(* IEC 61131-3 sources: JingjiangMoonbox/Application/Application/任务列表/CommTask/参数初始化 (part 2) *)

(* ---- KS_RstGrpParam_UnSave.st ---- *)
(*@CES
Name=KS_RstGrpParam_UnSave
Type=FunctionBlock
TypeGuid=6f9dac99-8de1-4efc-8465-68ac443b7d08
Guid=192eb973-c984-42d3-866b-81e626ce7a5f
HasDeclaration=True
HasImplementation=True
*)
{DECLARATION}
FUNCTION KS_RstGrpParam_UnSave : INT
VAR_INPUT
	i_pastStGrpParam_UnSave: POINTER TO ARRAY [1..2] OF StGrpParam_UnSave;
	i_pastStGrpParam_UnSave_RSV: POINTER TO ARRAY [1..2] OF StRSV_GrpParam_UnSave;
END_VAR
VAR
	iGrp: INT;
	iResult: INT;
	iT: INT;
END_VAR

{IMPLEMENTATION}
iResult:=0;

IF i_pastStGrpParam_UnSave<>0 AND i_pastStGrpParam_UnSave_RSV<>0 THEN
	FOR iGrp:=1 TO 2 BY 1 DO
		SysMemSet(ADR(i_pastStGrpParam_UnSave_RSV^[iGrp].abyRSV_StGrpParam_UnSave),
					0,
					SIZEOF(i_pastStGrpParam_UnSave_RSV^[iGrp].abyRSV_StGrpParam_UnSave));
		i_pastStGrpParam_UnSave^[iGrp].xCutterOnTop_Uw						:= TRUE;
		i_pastStGrpParam_UnSave^[iGrp].iDebugVelmpm_AxisA_Uw                := 100;
		i_pastStGrpParam_UnSave^[iGrp].iDebugGirthmm_AxisA_Uw               := 300;
		i_pastStGrpParam_UnSave^[iGrp].iDebugVelmpm_AxisB_Uw                := 100;
		i_pastStGrpParam_UnSave^[iGrp].iDebugGirthmm_AxisB_Uw               := 300;
		i_pastStGrpParam_UnSave^[iGrp].iDebugVelmpm_AxisA_Rw                := 100;
		i_pastStGrpParam_UnSave^[iGrp].iDebugGirthmm_AxisA_Rw               := 300;
		i_pastStGrpParam_UnSave^[iGrp].iDebugVelmpm_AxisB_Rw                := 100;
		i_pastStGrpParam_UnSave^[iGrp].iDebugGirthmm_AxisB_Rw               := 300;
		i_pastStGrpParam_UnSave^[iGrp].xMachineRev                          := FALSE;
		i_pastStGrpParam_UnSave^[iGrp].iPromptMsg                           := 0;
		i_pastStGrpParam_UnSave^[iGrp].iAlarm_TypeId                        := 0;
		i_pastStGrpParam_UnSave^[iGrp].iAlarm_UnitId                        := 0;
		i_pastStGrpParam_UnSave^[iGrp].iIdGSE                               := GSE_STOP;
		i_pastStGrpParam_UnSave^[iGrp].xFlag_Stop                           := TRUE;
		i_pastStGrpParam_UnSave^[iGrp].xFlag_PreStart                       := FALSE;
		i_pastStGrpParam_UnSave^[iGrp].xFlag_Ink                            := FALSE;
		i_pastStGrpParam_UnSave^[iGrp].xFlag_InkAccing                      := FALSE;
		i_pastStGrpParam_UnSave^[iGrp].xFlag_Tension                        := FALSE;
		i_pastStGrpParam_UnSave^[iGrp].xFlag_TensionDone                    := FALSE;
		i_pastStGrpParam_UnSave^[iGrp].xFlag_Print                          := FALSE;
		i_pastStGrpParam_UnSave^[iGrp].xFlag_Estop                          := FALSE;
		i_pastStGrpParam_UnSave^[iGrp].xFlag_AutoAcc                        := FALSE;
		i_pastStGrpParam_UnSave^[iGrp].xFlag_AutoDec                        := FALSE;
		i_pastStGrpParam_UnSave^[iGrp].xFlag_ManuAcc                        := FALSE;
		i_pastStGrpParam_UnSave^[iGrp].xFlag_ManuDec                        := FALSE;
		i_pastStGrpParam_UnSave^[iGrp].xFlag_Accing                         := FALSE;
		i_pastStGrpParam_UnSave^[iGrp].xFlag_Decing                         := FALSE;
		i_pastStGrpParam_UnSave^[iGrp].xFlag_EStoping                       := FALSE;
		i_pastStGrpParam_UnSave^[iGrp].xFlag_Stoping                        := FALSE;
		i_pastStGrpParam_UnSave^[iGrp].xFlag_GotoInking                     := FALSE;
		i_pastStGrpParam_UnSave^[iGrp].xFlag_InPressing                     := FALSE;
		i_pastStGrpParam_UnSave^[iGrp].xFlag_RollerPressDone                := FALSE;
		i_pastStGrpParam_UnSave^[iGrp].xFlag_InchRun                        := FALSE;
		i_pastStGrpParam_UnSave^[iGrp].xFlag_AllInchRun                     := FALSE;
		i_pastStGrpParam_UnSave^[iGrp].xFlag_AllPress                       := FALSE;
		i_pastStGrpParam_UnSave^[iGrp].xFlag_AllUnpress                     := FALSE;
		i_pastStGrpParam_UnSave^[iGrp].xFlag_RollerPressAtLeast1            := FALSE;
		i_pastStGrpParam_UnSave^[iGrp].axFlag_PrnLen_Alarm[1]                  := FALSE;
		i_pastStGrpParam_UnSave^[iGrp].axFlag_PrnLen_Alarm[2]                  := FALSE;
		i_pastStGrpParam_UnSave^[iGrp].axFlag_PrnLen_Alarm[3]                  := FALSE;
		i_pastStGrpParam_UnSave^[iGrp].xFlag_LinkageAxisAlarm               := FALSE;
		i_pastStGrpParam_UnSave^[iGrp].xFlag_TensionUnfinished              := FALSE;
		i_pastStGrpParam_UnSave^[iGrp].xFlag_VelTooHigh                     := FALSE;
		i_pastStGrpParam_UnSave^[iGrp].xFlag_PrestartTimeout                := FALSE;
		i_pastStGrpParam_UnSave^[iGrp].xFlag_KeepAlarming                   := FALSE;
		i_pastStGrpParam_UnSave^[iGrp].xFlag_ArrivedToTargetVel             := FALSE;
		i_pastStGrpParam_UnSave^[iGrp].xFlag_FilmAccDecDone                 := FALSE;
		i_pastStGrpParam_UnSave^[iGrp].xSlowStopTenEn                       := FALSE;
		i_pastStGrpParam_UnSave^[iGrp].xIsDebugMode_Machine                 := FALSE;
		i_pastStGrpParam_UnSave^[iGrp].uiFilmThickNess                      := 20;
		i_pastStGrpParam_UnSave^[iGrp].abyClrPrnLenCount_Rw[1]                 := 0;
		i_pastStGrpParam_UnSave^[iGrp].abyClrPrnLenCount_Rw[2]                 := 0;
		i_pastStGrpParam_UnSave^[iGrp].abyClrPrnLenCount_Rw[3]                 := 0;
		i_pastStGrpParam_UnSave^[iGrp].iTimeSec_AccDec_AllTheWay            := 0;
		i_pastStGrpParam_UnSave^[iGrp].rAccDecTime_ThisTime                 := 0;
		i_pastStGrpParam_UnSave^[iGrp].alrStdVol_Diam_Axis_Hmi[1]              := 0;
		i_pastStGrpParam_UnSave^[iGrp].alrStdVol_Diam_Axis_Hmi[2]              := 0;
		i_pastStGrpParam_UnSave^[iGrp].alrStdVol_Diam_Axis_Hmi[3]              := 0;
		i_pastStGrpParam_UnSave^[iGrp].alrStdVol_Diam_Axis_Hmi[4]              := 0;
		i_pastStGrpParam_UnSave^[iGrp].alrStdVol_Volt_Axis_Hmi[1]              := 0;
		i_pastStGrpParam_UnSave^[iGrp].alrStdVol_Volt_Axis_Hmi[2]              := 0;
		i_pastStGrpParam_UnSave^[iGrp].alrStdVol_Volt_Axis_Hmi[3]              := 0;
		i_pastStGrpParam_UnSave^[iGrp].alrStdVol_Volt_Axis_Hmi[4]              := 0;
		i_pastStGrpParam_UnSave^[iGrp].alrStdVol_Coef_Axis_Hmi[0]              := 0;
		i_pastStGrpParam_UnSave^[iGrp].alrStdVol_Coef_Axis_Hmi[1]              := 0;
		i_pastStGrpParam_UnSave^[iGrp].alrStdVol_Coef_Axis_Hmi[2]              := 0;
		i_pastStGrpParam_UnSave^[iGrp].alrStdVol_Coef_Axis_Hmi[3]              := 0;
		i_pastStGrpParam_UnSave^[iGrp].alrStdVol_Coef_Axis_Hmi[4]              := 0;
		i_pastStGrpParam_UnSave^[iGrp].rVel_Cur                             := 0;
		i_pastStGrpParam_UnSave^[iGrp].rVel_Film                            := 0;
		i_pastStGrpParam_UnSave^[iGrp].iSid_AxisA_Uw                        := 112;
		i_pastStGrpParam_UnSave^[iGrp].xStationOnline_AxisA_Uw              := FALSE;
		i_pastStGrpParam_UnSave^[iGrp].xMotRev_AxisA_Uw                     := FALSE;
		i_pastStGrpParam_UnSave^[iGrp].iSid_AxisB_Uw                        := 113;
		i_pastStGrpParam_UnSave^[iGrp].xStationOnline_AxisB_Uw              := FALSE;
		i_pastStGrpParam_UnSave^[iGrp].xMotRev_AxisB_Uw                     := FALSE;
		i_pastStGrpParam_UnSave^[iGrp].rAI_Uw                               := 0;
		i_pastStGrpParam_UnSave^[iGrp].rAI_Act_Uw                           := 0;
		i_pastStGrpParam_UnSave^[iGrp].rAI_HMI_Uw                           := 0;
		i_pastStGrpParam_UnSave^[iGrp].rAI_DiamMeasure_Uw                   := 0;
		i_pastStGrpParam_UnSave^[iGrp].arKpid_Current_Uw[1]                    := 20;
		i_pastStGrpParam_UnSave^[iGrp].arKpid_Current_Uw[2]                    := 50;
		i_pastStGrpParam_UnSave^[iGrp].arKpid_Current_Uw[3]                    := 50;
		i_pastStGrpParam_UnSave^[iGrp].arKpid_Current_Rw[1]                    := 0;
		i_pastStGrpParam_UnSave^[iGrp].arKpid_Current_Rw[2]                    := 0;
		i_pastStGrpParam_UnSave^[iGrp].arKpid_Current_Rw[3]                    := 0;
		i_pastStGrpParam_UnSave^[iGrp].rVel_PreDrv_Uw                       := 0;
		i_pastStGrpParam_UnSave^[iGrp].xReflectionSensorValid_Uw            := FALSE;
		i_pastStGrpParam_UnSave^[iGrp].xReflectSensorLoss_Uw                := FALSE;
		i_pastStGrpParam_UnSave^[iGrp].rDiam_NewVol_Uw                      := 400;
		i_pastStGrpParam_UnSave^[iGrp].rTowerThetaCur_Uw                    := 0;
		i_pastStGrpParam_UnSave^[iGrp].rFilmToTowerRollerDis_Uw             := 0;
		i_pastStGrpParam_UnSave^[iGrp].xFilmTouchRoller_Uw                  := FALSE;
		i_pastStGrpParam_UnSave^[iGrp].xSts_PreCutting_Uw                   := FALSE;
		i_pastStGrpParam_UnSave^[iGrp].rDebugCurVelmpmAxisA_Uw              := 0;
		i_pastStGrpParam_UnSave^[iGrp].rDebugCurVelrpmAxisA_Uw              := 0;
		i_pastStGrpParam_UnSave^[iGrp].rDebugCurVelmpmAxisB_Uw              := 0;
		i_pastStGrpParam_UnSave^[iGrp].rDebugCurVelrpmAxisB_Uw              := 0;
		i_pastStGrpParam_UnSave^[iGrp].rDeltaW_RPMIN_Uw                     := 0;
		i_pastStGrpParam_UnSave^[iGrp].xDebugMode_AbsEnc_Uw                 := FALSE;
		i_pastStGrpParam_UnSave^[iGrp].dwAbsEncSinglePos_Uw                 := 0;
		i_pastStGrpParam_UnSave^[iGrp].dwAbsEncSPos_Cur_Uw                  := 0;
		i_pastStGrpParam_UnSave^[iGrp].byEncodeValueWr_Uw                   := 0;
		i_pastStGrpParam_UnSave^[iGrp].rAIByAbsEnc_Cur_Uw                   := 0;
		i_pastStGrpParam_UnSave^[iGrp].xCutterOnTopFroDebug_Uw              := FALSE;
		i_pastStGrpParam_UnSave^[iGrp].xCurAxisAFroDebug_Uw                 := FALSE;
		i_pastStGrpParam_UnSave^[iGrp].xAlarmBell_Uw                        := FALSE;
		i_pastStGrpParam_UnSave^[iGrp].xIsDebug_DiaMeasure_Uw               := FALSE;
		i_pastStGrpParam_UnSave^[iGrp].byIsDebug_DiaMeasureArea_Uw          := 0;
		i_pastStGrpParam_UnSave^[iGrp].xIsDebuging_DiaMeasure_Uw            := FALSE;
		i_pastStGrpParam_UnSave^[iGrp].xCancelDebuging_DiaMeasure_Uw        := FALSE;
		i_pastStGrpParam_UnSave^[iGrp].byAxisDebugBit_Uw                    := 0;
		i_pastStGrpParam_UnSave^[iGrp].byAxisDebugBit_Uw_2                  := 0;
		i_pastStGrpParam_UnSave^[iGrp].xEnCodeErr_Uw                        := FALSE;
		i_pastStGrpParam_UnSave^[iGrp].xEnCodeErr_Rw                        := FALSE;
		i_pastStGrpParam_UnSave^[iGrp].rPi_Value_Uw                         := 0;
		i_pastStGrpParam_UnSave^[iGrp].rForwardStep_Uw                      := 0;
		i_pastStGrpParam_UnSave^[iGrp].xAxisAForeward_Uw                    := FALSE;
		i_pastStGrpParam_UnSave^[iGrp].xAxisBForeward_Uw                    := FALSE;
		i_pastStGrpParam_UnSave^[iGrp].rVelRPM_Cur_Uw                       := 0;
		i_pastStGrpParam_UnSave^[iGrp].rAxisAVelRPM_Cur_Uw                  := 0;
		i_pastStGrpParam_UnSave^[iGrp].rAxisBVelRPM_Cur_Uw                  := 0;
		i_pastStGrpParam_UnSave^[iGrp].xFlag_DiamCalc_ing_Uw                := FALSE;
		i_pastStGrpParam_UnSave^[iGrp].xFlag_DiamCalc_end_Uw                := FALSE;
		i_pastStGrpParam_UnSave^[iGrp].xFlag_DiamMeasure_end_Uw             := FALSE;
		i_pastStGrpParam_UnSave^[iGrp].xFlag_PreDrv_ing_Uw                  := FALSE;
		i_pastStGrpParam_UnSave^[iGrp].xFlag_PreDrv_end_Uw                  := FALSE;

		i_pastStGrpParam_UnSave^[iGrp].xFlag_Cut_end_Uw_UseInOtherPrg:= FALSE;
		i_pastStGrpParam_UnSave^[iGrp].xFlag_Cut_ing_Uw_UseInOtherPrg:= FALSE;
		i_pastStGrpParam_UnSave^[iGrp].xFlag_Cut_end_Uw:= TRUE;
		i_pastStGrpParam_UnSave^[iGrp].xFlag_Cut_ing_Uw:= FALSE;

		i_pastStGrpParam_UnSave^[iGrp].xFlag_VolDiamAlarm_Uw                := FALSE;
		i_pastStGrpParam_UnSave^[iGrp].rAI_DiamMeasure_HMI_Uw               := 0;
		i_pastStGrpParam_UnSave^[iGrp].xAITypeBtn_Uw                        := FALSE;
		i_pastStGrpParam_UnSave^[iGrp].iSid_AxisA_Rw                        := 114;
		i_pastStGrpParam_UnSave^[iGrp].xStationOnline_AxisA_Rw              := FALSE;
		i_pastStGrpParam_UnSave^[iGrp].xMotRev_AxisA_Rw                     := FALSE;
		i_pastStGrpParam_UnSave^[iGrp].iSid_AxisB_Rw                        := 115;
		i_pastStGrpParam_UnSave^[iGrp].xStationOnline_AxisB_Rw              := FALSE;
		i_pastStGrpParam_UnSave^[iGrp].xMotRev_AxisB_Rw                     := FALSE;
		i_pastStGrpParam_UnSave^[iGrp].rAI_Rw                               := 0;
		i_pastStGrpParam_UnSave^[iGrp].rAI_Act_Rw                           := 0;
		i_pastStGrpParam_UnSave^[iGrp].rAI_HMI_Rw                           := 0;
		i_pastStGrpParam_UnSave^[iGrp].rVel_PreDrv_Rw                       := 0;
		i_pastStGrpParam_UnSave^[iGrp].rDiam_NewVol_Rw                      := 0;
		i_pastStGrpParam_UnSave^[iGrp].rTaper_Rw                            := 0;
		i_pastStGrpParam_UnSave^[iGrp].xSts_PreCutting_Rw                   := FALSE;
		i_pastStGrpParam_UnSave^[iGrp].rDebugCurVelmpmAxisA_Rw              := 0;
		i_pastStGrpParam_UnSave^[iGrp].rDebugCurVelrpmAxisA_Rw              := 0;
		i_pastStGrpParam_UnSave^[iGrp].rDebugCurVelmpmAxisB_Rw              := 0;
		i_pastStGrpParam_UnSave^[iGrp].rDebugCurVelrpmAxisB_Rw              := 0;
		i_pastStGrpParam_UnSave^[iGrp].xDebugMode_AbsEnc_Rw                 := FALSE;
		i_pastStGrpParam_UnSave^[iGrp].dwAbsEncSinglePos_Rw                 := 0;
		i_pastStGrpParam_UnSave^[iGrp].dwAbsEncSPos_Cur_Rw                  := 0;
		i_pastStGrpParam_UnSave^[iGrp].byEncodeValueWr_Rw                   := 0;
		i_pastStGrpParam_UnSave^[iGrp].xCutterOnTopFroDebug_Rw              := FALSE;
		i_pastStGrpParam_UnSave^[iGrp].xCurAxisAFroDebug_Rw                 := FALSE;
		i_pastStGrpParam_UnSave^[iGrp].x6InchFroDebug_Rw                    := FALSE;
		i_pastStGrpParam_UnSave^[iGrp].xAlarmBell_Rw                        := FALSE;
		i_pastStGrpParam_UnSave^[iGrp].byAxisDebugBit_Rw                    := 0;
		i_pastStGrpParam_UnSave^[iGrp].rPi_Value_Rw                         := 0;
		i_pastStGrpParam_UnSave^[iGrp].rForwardStep_Rw                      := 0;
		i_pastStGrpParam_UnSave^[iGrp].xAxisAForeward_Rw                    := FALSE;
		i_pastStGrpParam_UnSave^[iGrp].xAxisBForeward_Rw                    := FALSE;
		i_pastStGrpParam_UnSave^[iGrp].rVelRPM_Cur_Rw                       := 0;
		i_pastStGrpParam_UnSave^[iGrp].rAxisAVelRPM_Cur_Rw                  := 0;
		i_pastStGrpParam_UnSave^[iGrp].rAxisBVelRPM_Cur_Rw                  := 0;
		i_pastStGrpParam_UnSave^[iGrp].xFlag_6Inch_Rw                       := FALSE;
		i_pastStGrpParam_UnSave^[iGrp].xFlag_PreDrv_ing_Rw                  := FALSE;
		i_pastStGrpParam_UnSave^[iGrp].xFlag_PreDrv_end_Rw                  := FALSE;
		i_pastStGrpParam_UnSave^[iGrp].xFlag_Cut_ing_Rw                     := FALSE;
		i_pastStGrpParam_UnSave^[iGrp].xFlag_Cut_end_Rw                     := FALSE;
		i_pastStGrpParam_UnSave^[iGrp].xAITypeBtn_Rw                        := FALSE;
		i_pastStGrpParam_UnSave^[iGrp].iSid_If                              := 120;
		i_pastStGrpParam_UnSave^[iGrp].xStationOnline_If                    := FALSE;
		i_pastStGrpParam_UnSave^[iGrp].xMotRev_If                           := FALSE;
		i_pastStGrpParam_UnSave^[iGrp].rAI_If                               := 0;
		i_pastStGrpParam_UnSave^[iGrp].rAI_Act_If                           := 0;
		i_pastStGrpParam_UnSave^[iGrp].rAI_HMI_If                           := 0;
		i_pastStGrpParam_UnSave^[iGrp].xInchBtn_If                          := FALSE;
		i_pastStGrpParam_UnSave^[iGrp].xRollerSts_If                        := FALSE;
		i_pastStGrpParam_UnSave^[iGrp].xRunEn_If                            := FALSE;
		i_pastStGrpParam_UnSave^[iGrp].rVel_Cur_If                          := 0;
		i_pastStGrpParam_UnSave^[iGrp].rPi_Value_If                         := 0;
		i_pastStGrpParam_UnSave^[iGrp].rForwardStep_If                      := 0;
		i_pastStGrpParam_UnSave^[iGrp].rUsingGirth_If                       := 0;
		i_pastStGrpParam_UnSave^[iGrp].xInching_If                          := FALSE;
		i_pastStGrpParam_UnSave^[iGrp].xAITypeBtn_if                        := FALSE;
		i_pastStGrpParam_UnSave^[iGrp].iSid_Of                              := 121;
		i_pastStGrpParam_UnSave^[iGrp].xStationOnline_Of                    := FALSE;
		i_pastStGrpParam_UnSave^[iGrp].xMotRev_Of                           := FALSE;
		i_pastStGrpParam_UnSave^[iGrp].rAI_Of                               := 0;
		i_pastStGrpParam_UnSave^[iGrp].rAI_Act_Of                           := 0;
		i_pastStGrpParam_UnSave^[iGrp].rAI_HMI_Of                           := 0;
		i_pastStGrpParam_UnSave^[iGrp].xInchBtn_Of                          := FALSE;
		i_pastStGrpParam_UnSave^[iGrp].xRollerSts_Of                        := FALSE;
		i_pastStGrpParam_UnSave^[iGrp].xRunEn_Of                            := FALSE;
		i_pastStGrpParam_UnSave^[iGrp].rVel_Cur_Of                          := 0;
		i_pastStGrpParam_UnSave^[iGrp].rPi_Value_Of                         := 0;
		i_pastStGrpParam_UnSave^[iGrp].rForwardStep_Of                      := 0;
		i_pastStGrpParam_UnSave^[iGrp].rUsingGirth_Of                       := 0;
		i_pastStGrpParam_UnSave^[iGrp].xInching_Of                          := FALSE;
		i_pastStGrpParam_UnSave^[iGrp].xAITypeBtn_Of                        := FALSE;
		i_pastStGrpParam_UnSave^[iGrp].sCurRecipeName_InUse                 := '';
		i_pastStGrpParam_UnSave^[iGrp].dwSTS_ALL                            := 0;
		i_pastStGrpParam_UnSave^[iGrp].xAutoAccDec_Hmi                      := FALSE;
		i_pastStGrpParam_UnSave^[iGrp].xFlag_IfOf_Ink                       := FALSE;
		i_pastStGrpParam_UnSave^[iGrp].xFlag_FastStoping                    := FALSE;
		i_pastStGrpParam_UnSave^[iGrp].rFinalVelocity                       := 0;
		i_pastStGrpParam_UnSave^[iGrp].xFlag_AutoMaticCutting_Uw            := FALSE;
		i_pastStGrpParam_UnSave^[iGrp].xFlag_AutoMaticCutting_rw            := FALSE;
		i_pastStGrpParam_UnSave^[iGrp].rAutoMaticCuttingLenth_CurMode_uw    := 0;
		i_pastStGrpParam_UnSave^[iGrp].rActRemainFilmLenth_Uw               := 0;
		i_pastStGrpParam_UnSave^[iGrp].rAutoMaticCuttingLenth_CurMode_Rw    := 0;
		i_pastStGrpParam_UnSave^[iGrp].xCurAxisDia_Uw_Wr                    := FALSE;
		i_pastStGrpParam_UnSave^[iGrp].xCurAxisDia_Rw_Wr                    := FALSE;
		i_pastStGrpParam_UnSave^[iGrp].rTaper_Cur_Uw                        := 0;
		i_pastStGrpParam_UnSave^[iGrp].rTaper_Cur_If                        := 0;
		i_pastStGrpParam_UnSave^[iGrp].rTaper_Cur_Of                        := 0;
		i_pastStGrpParam_UnSave^[iGrp].rTaperValueBegin_Hmi_Uw              := 0;
		i_pastStGrpParam_UnSave^[iGrp].rTaperValueEnd_Hmi_Uw                := 0;
		i_pastStGrpParam_UnSave^[iGrp].rTaperValueBegin_Hmi_Rw              := 0;
		i_pastStGrpParam_UnSave^[iGrp].rTaperValueEnd_Hmi_Rw                := 0;
		i_pastStGrpParam_UnSave^[iGrp].rTaperValueBegin_Hmi_If              := 0;
		i_pastStGrpParam_UnSave^[iGrp].rTaperValueEnd_Hmi_If                := 0;
		i_pastStGrpParam_UnSave^[iGrp].rTaperValueBegin_Hmi_Of              := 0;
		i_pastStGrpParam_UnSave^[iGrp].rTaperValueEnd_Hmi_Of                := 0;
		i_pastStGrpParam_UnSave^[iGrp].byTaperUnitConfirm_Uw                := 0;
		i_pastStGrpParam_UnSave^[iGrp].byTaperUnitConfirm_Rw                := 0;
		i_pastStGrpParam_UnSave^[iGrp].byTaperUnitConfirm_If                := 0;
		i_pastStGrpParam_UnSave^[iGrp].byTaperUnitConfirm_Of                := 0;
		i_pastStGrpParam_UnSave^[iGrp].rTaperValueCur_Hmi_If                := 0;
		i_pastStGrpParam_UnSave^[iGrp].rTaperValueCur_Hmi_of                := 0;
		i_pastStGrpParam_UnSave^[iGrp].rTaperValueCur_Hmi_Uw                := 0;
		i_pastStGrpParam_UnSave^[iGrp].rTaperValueCur_Hmi_Rw                := 0;
		i_pastStGrpParam_UnSave^[iGrp].rValue_DiaMeasure                    := 0;
		i_pastStGrpParam_UnSave^[iGrp].rVolt_CalcDiam_Used_Watch            := 0;
		i_pastStGrpParam_UnSave^[iGrp].rAO_Inverter_Uw_AxisA                := 0;
		i_pastStGrpParam_UnSave^[iGrp].rAO_Inverter_Uw_AxisB                := 0;
		i_pastStGrpParam_UnSave^[iGrp].rAO_Inverter_Rw_AxisA                := 0;
		i_pastStGrpParam_UnSave^[iGrp].rAO_Inverter_Rw_AxisB                := 0;
		i_pastStGrpParam_UnSave^[iGrp].xBtn_HorzPreRegister_Repeat          := FALSE;
		i_pastStGrpParam_UnSave^[iGrp].xBtn_HorzPreRegister_Setup           := FALSE;
		i_pastStGrpParam_UnSave^[iGrp].xSts_HorzPreRegister                 := FALSE;
		i_pastStGrpParam_UnSave^[iGrp].xMode_HorzPreRegister                := FALSE;
		i_pastStGrpParam_UnSave^[iGrp].xFlag_HorzPreRegister_All_end        := FALSE;
		i_pastStGrpParam_UnSave^[iGrp].xFlag_Home                           := FALSE;
		i_pastStGrpParam_UnSave^[iGrp].xFlag_Home_ing                       := FALSE;
		i_pastStGrpParam_UnSave^[iGrp].xFlag_Home_end                       := FALSE;
		i_pastStGrpParam_UnSave^[iGrp].xFlag_ConfirmPreRegHomePos           := FALSE;
		i_pastStGrpParam_UnSave^[iGrp].xFlag_ConfirmPreRegHomePos_ing       := FALSE;
		i_pastStGrpParam_UnSave^[iGrp].xFlag_ConfirmPreRegHomePos_end       := FALSE;
		i_pastStGrpParam_UnSave^[iGrp].xFlag_PreRegister                    := FALSE;
		i_pastStGrpParam_UnSave^[iGrp].xFlag_PreRegister_ing                := FALSE;
		i_pastStGrpParam_UnSave^[iGrp].xFlag_PreRegister_end                := FALSE;
		i_pastStGrpParam_UnSave^[iGrp].xFlag_PhaseRestore                   := FALSE;
		i_pastStGrpParam_UnSave^[iGrp].xFlag_PhaseRestore_ing               := FALSE;
		i_pastStGrpParam_UnSave^[iGrp].xFlag_PhaseRestore_end               := FALSE;
		i_pastStGrpParam_UnSave^[iGrp].xBtn_Home                            := FALSE;
		i_pastStGrpParam_UnSave^[iGrp].xBtn_ConfirmPreRegHomePos            := FALSE;
		i_pastStGrpParam_UnSave^[iGrp].xBtn_PreRegister                     := FALSE;
		i_pastStGrpParam_UnSave^[iGrp].xBtn_PhaseSave                       := FALSE;
		i_pastStGrpParam_UnSave^[iGrp].xBtn_PhaseRestore                    := FALSE;
		i_pastStGrpParam_UnSave^[iGrp].xFlag_MotionParamInitialized         := FALSE;
		i_pastStGrpParam_UnSave^[iGrp].xFlag_AccDecStop                     := FALSE;
		i_pastStGrpParam_UnSave^[iGrp].xNetOffline_CENTRAL                  := FALSE;
		i_pastStGrpParam_UnSave^[iGrp].xAxisAlarm_CENTRAL                   := FALSE;
		i_pastStGrpParam_UnSave^[iGrp].xPosDeviationAlarm_CENTRAL           := FALSE;
		i_pastStGrpParam_UnSave^[iGrp].xNetOffline_CENTRAL2                 := FALSE;
		i_pastStGrpParam_UnSave^[iGrp].xAxisAlarm_CENTRAL2                  := FALSE;
		i_pastStGrpParam_UnSave^[iGrp].xPosDeviationAlarm_CENTRAL2          := FALSE;
		i_pastStGrpParam_UnSave^[iGrp].xNetOffline_IF                       := FALSE;
		i_pastStGrpParam_UnSave^[iGrp].xAxisAlarm_IF                        := FALSE;
		i_pastStGrpParam_UnSave^[iGrp].xPosDeviationAlarm_IF                := FALSE;
		i_pastStGrpParam_UnSave^[iGrp].xNetOffline_OF                       := FALSE;
		i_pastStGrpParam_UnSave^[iGrp].xAxisAlarm_OF                        := FALSE;
		i_pastStGrpParam_UnSave^[iGrp].xPosDeviationAlarm_OF                := FALSE;
		i_pastStGrpParam_UnSave^[iGrp].xNetOffline_UW_A                     := FALSE;
		i_pastStGrpParam_UnSave^[iGrp].xAxisAlarm_UW_A                      := FALSE;
		i_pastStGrpParam_UnSave^[iGrp].xPosDeviationAlarm_UW_A              := FALSE;
		i_pastStGrpParam_UnSave^[iGrp].xNetOffline_UW_B                     := FALSE;
		i_pastStGrpParam_UnSave^[iGrp].xAxisAlarm_UW_B                      := FALSE;
		i_pastStGrpParam_UnSave^[iGrp].xPosDeviationAlarm_UW_B              := FALSE;
		i_pastStGrpParam_UnSave^[iGrp].xNetOffline_RW_A                     := FALSE;
		i_pastStGrpParam_UnSave^[iGrp].xAxisAlarm_RW_A                      := FALSE;
		i_pastStGrpParam_UnSave^[iGrp].xPosDeviationAlarm_RW_A              := FALSE;
		i_pastStGrpParam_UnSave^[iGrp].xNetOffline_RW_B                     := FALSE;
		i_pastStGrpParam_UnSave^[iGrp].xAxisAlarm_RW_B                      := FALSE;
		i_pastStGrpParam_UnSave^[iGrp].xPosDeviationAlarm_RW_B              := FALSE;
		i_pastStGrpParam_UnSave^[iGrp].dwAlarmDetail_CENTRAL                := 0;
		i_pastStGrpParam_UnSave^[iGrp].dwAlarmDetail_CENTRAL2               := 0;
		i_pastStGrpParam_UnSave^[iGrp].dwAlarmDetail_IF                     := 0;
		i_pastStGrpParam_UnSave^[iGrp].dwAlarmDetail_OF                     := 0;
		i_pastStGrpParam_UnSave^[iGrp].dwAlarmDetail_UW_A                   := 0;
		i_pastStGrpParam_UnSave^[iGrp].dwAlarmDetail_UW_B                   := 0;
		i_pastStGrpParam_UnSave^[iGrp].dwAlarmDetail_RW_A                   := 0;
		i_pastStGrpParam_UnSave^[iGrp].dwAlarmDetail_RW_B                   := 0;
		i_pastStGrpParam_UnSave^[iGrp].xValid_CentralDrum                   := FALSE;
		i_pastStGrpParam_UnSave^[iGrp].iSid_CentralDrum                     := 16;
		i_pastStGrpParam_UnSave^[iGrp].xStationOnline_CentralDrum           := FALSE;
		i_pastStGrpParam_UnSave^[iGrp].xMotRev_CentralDrum                  := FALSE;
		i_pastStGrpParam_UnSave^[iGrp].rAxisVel_CentralDrum                 := 0;
		i_pastStGrpParam_UnSave^[iGrp].xPrintInching                        := FALSE;
		i_pastStGrpParam_UnSave^[iGrp].rVel_Inching_Print                   := 5;
		i_pastStGrpParam_UnSave^[iGrp].xTapPosition_Breaking                := FALSE;
		i_pastStGrpParam_UnSave^[iGrp].xTapPosition_UniformInk              := FALSE;
		i_pastStGrpParam_UnSave^[iGrp].xTapPosition_Printing                := FALSE;
		i_pastStGrpParam_UnSave^[iGrp].wEn_UwRw_IfOf_Center                 := 0;
		SysMemSet(ADR(i_pastStGrpParam_UnSave^[iGrp].aiMotionStep_AllStation ),
				0,
				SIZEOF(i_pastStGrpParam_UnSave^[iGrp].aiMotionStep_AllStation ));

		i_pastStGrpParam_UnSave^[iGrp].stStTimeSet_DnCut_UpCut_Uw_Hmi.iDelayMsec_CutterHolder:= 0;
		i_pastStGrpParam_UnSave^[iGrp].stStTimeSet_DnCut_UpCut_Uw_Hmi.iDelayMsec_CutOffKnifeCylinder:= 0;
		i_pastStGrpParam_UnSave^[iGrp].stStTimeSet_DnCut_UpCut_Uw_Hmi.iDelayMsec_RollerCylinder:= 0;
		i_pastStGrpParam_UnSave^[iGrp].stStTimeSet_DnCut_UpCut_Uw_Hmi.uiMM_Roller2GummedTape:= 0;
		i_pastStGrpParam_UnSave^[iGrp].stStTimeSet_DnCut_UpCut_Uw_Hmi.uiMM_Roller2CutOfKnife:= 0;
		i_pastStGrpParam_UnSave^[iGrp].stStTimeSet_DnCut_UpCut_Uw_Hmi.uiMM_CutOfKnife2GummedTape:= 0;
		i_pastStGrpParam_UnSave^[iGrp].stStTimeSet_DnCut_UpCut_Uw_Hmi.iStepVariation4ChangeTime:= 0;

		i_pastStGrpParam_UnSave^[iGrp].stStTimeSet_DnCut_UpCut_Rw_Hmi.iDelayMsec_CutterHolder:= 0;
		i_pastStGrpParam_UnSave^[iGrp].stStTimeSet_DnCut_UpCut_Rw_Hmi.iDelayMsec_CutOffKnifeCylinder:= 0;
		i_pastStGrpParam_UnSave^[iGrp].stStTimeSet_DnCut_UpCut_Rw_Hmi.iDelayMsec_RollerCylinder:= 0;
		i_pastStGrpParam_UnSave^[iGrp].stStTimeSet_DnCut_UpCut_Rw_Hmi.uiMM_Roller2GummedTape:= 0;
		i_pastStGrpParam_UnSave^[iGrp].stStTimeSet_DnCut_UpCut_Rw_Hmi.uiMM_Roller2CutOfKnife:= 0;
		i_pastStGrpParam_UnSave^[iGrp].stStTimeSet_DnCut_UpCut_Rw_Hmi.uiMM_CutOfKnife2GummedTape:= 0;
		i_pastStGrpParam_UnSave^[iGrp].stStTimeSet_DnCut_UpCut_Rw_Hmi.iStepVariation4ChangeTime:= 0;

		i_pastStGrpParam_UnSave^[iGrp].xPseudoRandomEn:= FALSE;
		i_pastStGrpParam_UnSave^[iGrp].byPseudoRandomId:= 1;
		i_pastStGrpParam_UnSave^[iGrp].aiTestPseudoRandom_Kp[1]:= 10;
		i_pastStGrpParam_UnSave^[iGrp].aiTestPseudoRandom_Kp[2]:= 15;
		i_pastStGrpParam_UnSave^[iGrp].aiTestPseudoRandom_Kp[3]:= 20;
		i_pastStGrpParam_UnSave^[iGrp].aiTestPseudoRandom_Kd[1]:= 20;
		i_pastStGrpParam_UnSave^[iGrp].aiTestPseudoRandom_Kd[2]:= 35;
		i_pastStGrpParam_UnSave^[iGrp].aiTestPseudoRandom_Kd[3]:= 40;
		i_pastStGrpParam_UnSave^[iGrp].xPseudoRandomTsting:= FALSE;
		i_pastStGrpParam_UnSave^[iGrp].xLinkage_IfOf_Ink:=FALSE;(*2022.4.9.235740*)
		i_pastStGrpParam_UnSave^[iGrp].xCurAxisDia_Uw_Wr:= FALSE;(*2022.4.9.235740*)
		i_pastStGrpParam_UnSave^[iGrp].xCurAxisDia_Rw_Wr:= FALSE;(*2022.4.9.235740*)
		(*2024.01.19.132742*)
		i_pastStGrpParam_UnSave^[iGrp].xFlag_Cut_end_Uw_UseInOtherPrg:=FALSE;
		i_pastStGrpParam_UnSave^[iGrp].xFlag_Cut_end_Rw_UseInOtherPrg:=FALSE;
		i_pastStGrpParam_UnSave^[iGrp].xFlag_Follow_1U_V_UwCut:= FALSE;
		i_pastStGrpParam_UnSave^[iGrp].xKeepAlarm_NoMaterial:= FALSE;

		i_pastStGrpParam_UnSave^[iGrp].xKnob_6Inch_Rw:= FALSE;
		i_pastStGrpParam_UnSave^[iGrp].x6InchFroDebug_Rw		:=FALSE;(*收料6寸标志|用于调试*)
		i_pastStGrpParam_UnSave^[iGrp].xWillAutoMaticPreCut_Uw:= FALSE;
		i_pastStGrpParam_UnSave^[iGrp].rAxisAFreq_Uw:= 0;
		i_pastStGrpParam_UnSave^[iGrp].rAxisBFreq_Uw:= 0;
		i_pastStGrpParam_UnSave^[iGrp].rAxisAFreq_Rw:= 0;
		i_pastStGrpParam_UnSave^[iGrp].rAxisBFreq_Rw:= 0;
		i_pastStGrpParam_UnSave^[iGrp].rWuCompensate_Uw:= 0;
		i_pastStGrpParam_UnSave^[iGrp].rWuCompensate_Rw:= 0;
		i_pastStGrpParam_UnSave^[iGrp].rWuCompensate_Act_Uw:= 0;
		i_pastStGrpParam_UnSave^[iGrp].rWuCompensate_Act_Rw:= 0;
		i_pastStGrpParam_UnSave^[iGrp].xEn_Disturbance_If:= FALSE;
		i_pastStGrpParam_UnSave^[iGrp].xEn_Disturbance_Of:= FALSE;
		i_pastStGrpParam_UnSave^[iGrp].rFreq_Disturbance_If:= 1;
		i_pastStGrpParam_UnSave^[iGrp].rAmplitude_Disturbance_If:= 1;
		i_pastStGrpParam_UnSave^[iGrp].uiTotalTime_Disturbance_If:= 0;
		i_pastStGrpParam_UnSave^[iGrp].xOuting_sin_If:= FALSE;
		i_pastStGrpParam_UnSave^[iGrp].rResult_sin_If:= 0;
		i_pastStGrpParam_UnSave^[iGrp].rFreq_Disturbance_Of:= 1;
		i_pastStGrpParam_UnSave^[iGrp].rAmplitude_Disturbance_Of:= 1;
		i_pastStGrpParam_UnSave^[iGrp].uiTotalTime_Disturbance_Of:= 0;
		i_pastStGrpParam_UnSave^[iGrp].xOuting_sin_Of:= FALSE;
		i_pastStGrpParam_UnSave^[iGrp].rResult_sin_Of:= 0;

		i_pastStGrpParam_UnSave^[iGrp].byPseudoRandomRoundTimes_Cur:= 0;

		i_pastStGrpParam_UnSave^[iGrp].xFlagFollow1U_AccDecing:= FALSE;

		i_pastStGrpParam_UnSave^[iGrp].xEnaTestARC_Ink:= FALSE;
		i_pastStGrpParam_UnSave^[iGrp].rAcceleration_Max:= 0;
		i_pastStGrpParam_UnSave^[iGrp].rAcceleration_Cur:= 0;

		i_pastStGrpParam_UnSave^[iGrp].byGrpAxisNum_Pu	:= 0;

		SysMemSet(ADR(i_pastStGrpParam_UnSave^[iGrp].abyGrpAxisList),0,SIZEOF(i_pastStGrpParam_UnSave^[iGrp].abyGrpAxisList));

		SysMemSet(ADR(i_pastStGrpParam_UnSave^[iGrp].abyGrpArcAxisList),0,SIZEOF(i_pastStGrpParam_UnSave^[iGrp].abyGrpArcAxisList));
		FOR iT:=1 TO MAX_UNIT_NUM BY 1 DO
			i_pastStGrpParam_UnSave^[iGrp].abyAxisList_CoatingPrn[iT]:= gc_byInvisCoatingPrnAxisIdx;
		END_FOR
		i_pastStGrpParam_UnSave^[iGrp].byAxisNum_CoatingPrn		:= 0(*BYTE*);(*涂布总轴数|*)
		i_pastStGrpParam_UnSave_RSV^[iGrp].xSwitch_GrpInkEn:=FALSE;
	END_FOR
	iResult:=1;
ELSE
	iResult:=-1;
END_IF

(* ---- KS_RstSysParam.st ---- *)
(*@CES
Name=KS_RstSysParam
Type=FunctionBlock
TypeGuid=6f9dac99-8de1-4efc-8465-68ac443b7d08
Guid=f9e1f4e0-8736-47b6-9a7b-51fe01553e23
HasDeclaration=True
HasImplementation=True
*)
{DECLARATION}
FUNCTION KS_RstSysParam : INT
VAR_INPUT
	i_pstStSysParam: POINTER TO StSysParam;
	i_xResetAllParam: BOOL;(*全部参数初始化*)
END_VAR
VAR
	iResult: INT;
	iUnit:INT;
END_VAR

{IMPLEMENTATION}
iResult:= 0;
IF i_pstStSysParam<>0 THEN
	IF i_xResetAllParam THEN
		KS_RstSysParam_Save(ADR(i_pstStSysParam^.stStSysParam_Save),
				ADR(i_pstStSysParam^.stStRSV_SysParam_Save),
	(*2026.5.28.150112增加预套准结构初始化*)
				g_pstStMechanicalParam_01,
				g_pstStMechanicalParam_02,
				g_pstStMechanicalParam_03,
				g_pstStMechanicalParam_05);
		KS_RstGrpParam_Save(ADR(i_pstStSysParam^.astStGrpParam_Save),
				ADR(i_pstStSysParam^.astStRSV_GrpParam_Save));
		KS_RstUnitParam_Save(i_pstStSysParam,
				ADR(i_pstStSysParam^.astStUnitParam_Save),
				ADR(i_pstStSysParam^.astStRSV_UnitParam_Save));
	ELSE
		KS_RstSysParam_UnSave(ADR(i_pstStSysParam^.stStSysParam_UnSave),
				ADR(i_pstStSysParam^.stStRSV_SysParam_UnSave));
		KS_RstGrpParam_UnSave(ADR(i_pstStSysParam^.astStGrpParam_UnSave),
				ADR(i_pstStSysParam^.astStRSV_GrpParam_UnSave));
		KS_RstUnitParam_UnSave(ADR(i_pstStSysParam^.astStUnitParam_UnSave),
				ADR(i_pstStSysParam^.astStRSV_UnitParam_UnSave));

	END_IF
	(*再清除一些原来保持的东西@2026.06.03.194958+ by liu.yt*)
	IF i_pstStSysParam<>0 THEN
		FOR iUnit:=1 TO MAX_UNIT_NUM BY 1 DO
			(*初始化为纵横向手动*)
			i_pstStSysParam^.astStUnitParam_Save[iUnit].dwFlag_Sts.0:= FALSE;
			i_pstStSysParam^.astStUnitParam_Save[iUnit].dwFlag_Sts.1:= FALSE;
		END_FOR
	END_IF

	iResult:= 1;
ELSE
	iResult:= -1;
END_IF
KS_RstSysParam:= iResult;

(* ---- KS_RstSysParam_Save.st ---- *)
(*@CES
Name=KS_RstSysParam_Save
Type=FunctionBlock
TypeGuid=6f9dac99-8de1-4efc-8465-68ac443b7d08
Guid=8442070d-5efa-4f31-a934-f12a469761f6
HasDeclaration=True
HasImplementation=True
*)
{DECLARATION}
FUNCTION KS_RstSysParam_Save : INT
VAR_INPUT
	i_pstStSysParam_Save: POINTER TO StSysParam_Save;
	i_pstStSysParam_Save_RSV: POINTER TO StRSV_SysParam_Save;

	i_pstStMechanicalParam_01: POINTER TO StMechanicalParam_01; (* 机械结构1| *)
	i_pstStMechanicalParam_02: POINTER TO StMechanicalParam_02; (* 机械结构2| *)
	i_pstStMechanicalParam_03: POINTER TO StMechanicalParam_03; (* 机械结构3| *)
	i_pstStMechanicalParam_05: POINTER TO StMechanicalParam_05; (* 机械结构5| *)(*2023.09.21.150812 同步*)

END_VAR
VAR
	iResult: INT;
END_VAR

{IMPLEMENTATION}
iResult:=0;

IF i_pstStSysParam_Save<>0 AND i_pstStSysParam_Save_RSV<>0 THEN
	SysMemSet(ADR(i_pstStSysParam_Save_RSV^.abyRSV_SysParam_Save),
				0,
				SIZEOF(i_pstStSysParam_Save_RSV^.abyRSV_SysParam_Save));
	i_pstStSysParam_Save^.dwFileVersion						:= 16#20250628;
	i_pstStSysParam_Save^.iCustomerId                       := 0;
	i_pstStSysParam_Save^.dwEquipmentProf                   := 0;
	i_pstStSysParam_Save^.iUnitMaxNum                       := 9;
	i_pstStSysParam_Save^.iCurveViewMaxRange                := 100;
	i_pstStSysParam_Save^.iTitleTextHeight                  := 16;
	i_pstStSysParam_Save^.iEntryTextHeight                  := 12;
	i_pstStSysParam_Save^.iLabelTextHeight                  := 12;
	i_pstStSysParam_Save^.iButtonTextHeight                 := 10;
	i_pstStSysParam_Save^.iMessageTextHeight                := 18;
	i_pstStSysParam_Save^.iRsvdTextHeight                   := 10;
	i_pstStSysParam_Save^.byLanguageId                      := 1;
	i_pstStSysParam_Save^.byMinutes_ScrSaver                := 3;
	i_pstStSysParam_Save^.iPointDensity_RS                  := 4;
	i_pstStSysParam_Save^.wCtlFlag_IndependentSettings      := 0;
(*	i_pstStSysParam_Save^.dwControlComplexBits              := 0;*)
	i_pstStSysParam_Save^.xFlag_CancelSafetyGrate			:= FALSE;
	i_pstStSysParam_Save^.xSwitch_ArcTest_V					:= TRUE;
	i_pstStSysParam_Save^.xSwitch_ArcTest_H					:= TRUE;
	i_pstStSysParam_Save^.xAllowLinkageChangeInRunning		:= FALSE;
	i_pstStSysParam_Save^.xChangLinkageStsWhenPrint			:= FALSE;

//2026.5.14.091013
//	i_pstStSysParam_Save^.astStMechanicalParamBuf           := 1;
	i_pstStSysParam_Save^.dwCtlSwitchRef                    := 0;
	i_pstStSysParam_Save^.byHorzCtlMode                   := 1;
	i_pstStSysParam_Save^.rStepDrivePosPPulse               := 0.0002;
	i_pstStSysParam_Save^.iStepDrivePulsePRev               := 6000;
	i_pstStSysParam_Save^.iStepDriveSa_Vel                  := 10;
	i_pstStSysParam_Save^.iStepDrivePreReg_Vel              := 50;
	i_pstStSysParam_Save^.iStepDriveManu_Vel                := 20;
	i_pstStSysParam_Save^.iStepDriveAuto_Vel                := 20;
	i_pstStSysParam_Save^.iStepDriveAccTime                 := 50;
	i_pstStSysParam_Save^.iStepDriveManu_Vel_Fast           := 40;
	i_pstStSysParam_Save^.byOverPercent_RatedRpm            := 10;
	i_pstStSysParam_Save^.rCurrent_Limit                    := 10;
	i_pstStSysParam_Save^.xWorkMode_Inch                    := FALSE;
	i_pstStSysParam_Save^.rHorCtl_PosPPulse                 := 0.000635;
	i_pstStSysParam_Save^.diHorCtl_PulsePRev                := 131072;
	i_pstStSysParam_Save^.rHorCtl_PreReg_Vel                := 2;
	i_pstStSysParam_Save^.rHorCtl_Manu_Vel                  := 0.5;
	i_pstStSysParam_Save^.rHorCtl_Manu_Vel_Fast             := 1;
	i_pstStSysParam_Save^.rHorCtl_Auto_Vel                  := 0.5;
	i_pstStSysParam_Save^.iHorCtl_Num                       := 60;
	i_pstStSysParam_Save^.iHorCtl_Den                       := 1;
	i_pstStSysParam_Save^.rHorCtl_Pitch                     := 5;
	i_pstStSysParam_Save^.iHorCtl_AccDecTime                := 10;
	i_pstStSysParam_Save^.diTimeHold_Prestart               := 3000;
	i_pstStSysParam_Save^.diTimeHold_Uw_Diam                := 3000;
	i_pstStSysParam_Save^.diTimeHold_Rw_Diam                := 3000;
	i_pstStSysParam_Save^.diTimeHold_Rw_Prnlength           := 3000;
	i_pstStSysParam_Save^.byHotBlowerStopDelayTime          := 0;
	i_pstStSysParam_Save^.byHeatingOutWay_III               := 1;
	i_pstStSysParam_Save^.iTimeOut_Slave_485_Inverter       := 3;
	i_pstStSysParam_Save^.iCofe_TempCtl_30                  := 30;
	i_pstStSysParam_Save^.iCofe_TempCtl_30_10               := 40;
	i_pstStSysParam_Save^.iCofe_TempCtl_10_5                := 50;
	i_pstStSysParam_Save^.iCofe_TempCtl_5                   := 60;
	i_pstStSysParam_Save^.iTime_Thres_Water                 := 150;
	i_pstStSysParam_Save^.byHeatingMode                     := 1;
	i_pstStSysParam_Save^.byOverTempValue                   := 150;
	i_pstStSysParam_Save^.byEn_ExtraFun_485                 := 16#0;
	i_pstStSysParam_Save^.iPidAlgorithm_Threshold           := 2;
	i_pstStSysParam_Save^.iMaxOutValue                      := 150;
	i_pstStSysParam_Save^.rKp                               := 10;
	i_pstStSysParam_Save^.rKi                               := 10;
	i_pstStSysParam_Save^.rKd                               := 300;
	i_pstStSysParam_Save^.uiCtrolCycle_Ms                   := 6000;
	i_pstStSysParam_Save^.iWaterValue_Threshold             := 60;
	i_pstStSysParam_Save^.iTempAcc_Threshold                := 20;
	i_pstStSysParam_Save^.iDecSV_PV_Threshold               := 10;
	i_pstStSysParam_Save^.xEn_HeatOff_AfterStop             := FALSE;
	i_pstStSysParam_Save^.xEn_HeatAirOff_AfterStop          := FALSE;
	i_pstStSysParam_Save^.rDelayOff_HotAir                  := 0;
	i_pstStSysParam_Save^.iDebugStep                        := 0;
	i_pstStSysParam_Save^.dwSwitch                          := 0;
//	i_pstStSysParam_Save^.byFakeThreshold_V                 := 50;
//	i_pstStSysParam_Save^.byFakeThreshold_H                 := 50;
//2026.5.29.185244补漏初始化
	i_pstStSysParam_Save^.xUnitPressOneBtn			:= FALSE;
	i_pstStSysParam_Save^.xAllPressOneBtn			:= FALSE;
	i_pstStSysParam_Save^.xPreCutOneBtn_Rw			:= FALSE;
	i_pstStSysParam_Save^.xPreCutOneBtn_Uw			:= FALSE;
	i_pstStSysParam_Save^.xTypeGetInitDiam:= TRUE;

	i_pstStSysParam_Save^.uiMaxDia:= 800;
	i_pstStSysParam_Save^.uiInitDiam_Uw:= 350;
	i_pstStSysParam_Save^.uiInitDiam_Rw:= 350;
	i_pstStSysParam_Save^.byCouplingType:= 0;

	(*新增加参数|wang.nt|2025.08.07.143540*)
	i_pstStSysParam_Save^.wMachineArchitectureRef									 :=0	;(*机器架构描述*)
	i_pstStSysParam_Save^.iPromptMsgId												 :=0	;(*提示信息ID（报警代码）*)
	i_pstStSysParam_Save^.byCheckTimeToTips_BrakeResistance							 :=1	;(*制动电阻访问超限提示时间*)
	i_pstStSysParam_Save^.byCheckTimeToEStop_BrakeResistance						:=4	;(*制动电阻访问超限急停时间*)
	i_pstStSysParam_Save^.byAccessTimes_BrakeResistance								 :=40	;(*制动电阻报警限制*)
	i_pstStSysParam_Save^.byAlarmHold_VOL_Uw										:=3	;(*放料没料响应时间*)
	i_pstStSysParam_Save^.byAlarmHold_PrnLength										 :=3	;(*收料印长报警响应时间*)
	i_pstStSysParam_Save^.rOpenThr_Ele												 :=0.9	;(*电加热开启*)
	i_pstStSysParam_Save^.rCloseThr_Ele												 :=0	;(*电加热关闭*)
	i_pstStSysParam_Save^.rDealValue_Water											 :=0.2	;(*水加热死区*)
	i_pstStSysParam_Save^.diStepDriveDebugPulse										 :=60000	;(*测试脉冲数*)
	i_pstStSysParam_Save^.iStepDriveDebugNum										:=1	;(*测试色组号*)
	i_pstStSysParam_Save^.rHz_MainExhaust_ManuallySet								 :=20	;(*主排风设定频率*)
	i_pstStSysParam_Save^.byFreq_I_ExhaustAir										 :=10	;(*排风一档频率*)
	i_pstStSysParam_Save^.byFreq_II_ExhaustAir										 :=20	;(*排风二档频率*)
	i_pstStSysParam_Save^.byFreq_III_ExhaustAir										 :=30	;(*排风三档频率*)
	(*9905界面参数*)
	i_pstStSysParam_Save^.byPseudoRandomRoundTimes									:=2		;
	i_pstStSysParam_Save^.rPseudoRandomAmplitude									:=0.03	;
	i_pstStSysParam_Save^.rCompensateGirthWhenAccing_If								:=0		;
	i_pstStSysParam_Save^.rCompensateGirthWhenAccing_Of								:=0		;
	i_pstStSysParam_Save^.iCustomerLogoOffsetX										:=-50	;
	i_pstStSysParam_Save^.byGuardrialColor_R										:=220	;
	i_pstStSysParam_Save^.byGuardrialColor_G										:=0		;
	i_pstStSysParam_Save^.byGuardrialColor_B										:=0		;
	i_pstStSysParam_Save^.iLedFuncId												:=0		;
	i_pstStSysParam_Save^.wRunningTime_Day											:=0		;
	i_pstStSysParam_Save^.byRunningTime_Hour										:=0		;
	i_pstStSysParam_Save^.byRunningTime_Min											:=0		;
	i_pstStSysParam_Save^.byRunningTime_Sec											:=0		;
	i_pstStSysParam_Save^.byArcIntensity_W											:=20		;
	i_pstStSysParam_Save^.byArcIntensity_M											:=15		;
	i_pstStSysParam_Save^.byArcIntensity_S											:=10		;
//2026.5.8.160718增加调整强度切换
	i_pstStSysParam_Save^.byArcIntensity											:=1		;

	i_pstStSysParam_Save^.byMotorOverTempValue_UseEncTemp							:=110		;
	i_pstStSysParam_Save^.byRemainSpaceNum_PTCTL									:=5		;
	i_pstStSysParam_Save^.rSpeed_SCoeff_Type789										:=2.0/3.0	;
	i_pstStSysParam_Save^.byMaxPulseOut_16dIO										:=3		;
	i_pstStSysParam_Save^.bySysSamplePrecision										:=2		;
	i_pstStSysParam_Save^.byArcAdjValueDealType										:=1		;
	i_pstStSysParam_Save^.byArcErrLimitToCtl_P										:=8		;
	i_pstStSysParam_Save^.byArcErrLimitToCtl_I 										:=1		;
	i_pstStSysParam_Save^.byMaxPulseOut_Module										:=15	;
	i_pstStSysParam_Save^.byArcFineSampleType										:=0		;
	i_pstStSysParam_Save^.byArcPidGetType 											:=0		;
	i_pstStSysParam_Save^.rFilmLenth_Eyes											:=1.5	;
	i_pstStSysParam_Save^.uiArcSysDelayTime_ms           							:=100	;
	i_pstStSysParam_Save^.byParamIndex_Huang										:=9		;
	i_pstStSysParam_Save^.uiControllerVel_Huang										:=0		;
	i_pstStSysParam_Save^.byDeCoupleArcNum											:=5		;
	i_pstStSysParam_Save^.xUseGc_PID_2025											:=TRUE	;(*2025.1.15.175536+*)
	i_pstStSysParam_Save^.byKadj_SetType											:= 0	;
	(*2025.8.19.211325增加*)
	i_pstStSysParam_Save^.byTypeFollow_Arc:= 0;(*先按照保持的处理*)
	i_pstStSysParam_Save^.byParamIndex_Huang:= 9;
	i_pstStSysParam_Save^.uiControllerVel_Huang:= 0;

	i_pstStSysParam_Save^.xInitArcErr_AjdImmediately:= TRUE;
	i_pstStSysParam_Save^.byUseArcAccOrDecCompensate:= 0;(*柔印先默认=0，不适用加速补偿*)

	i_pstStSysParam_Save^.xAutoSetArcCtlWay := TRUE;
	i_pstStSysParam_Save^.iUid:= 2;//2025.08.23.200449+
//2026.05.27.214505
	i_pstStSysParam_Save^.uiMaxVel_UseCalcAcc:= 100;

//2026.5.28.145220增加机械参数初始化
	IF i_pstStMechanicalParam_01<>0 THEN
		i_pstStMechanicalParam_01^.lrA			:= 90;(*LREAL*)
		i_pstStMechanicalParam_01^.lrD1			:= 100;(*LREAL*)
		i_pstStMechanicalParam_01^.lrD2			:= 100;(*LREAL*)
		i_pstStMechanicalParam_01^.lrD3			:= 100;(*LREAL*)
		i_pstStMechanicalParam_01^.lrDR			:= 135;(*LREAL*)
		i_pstStMechanicalParam_01^.lrL1			:= 225;(*LREAL*)
		i_pstStMechanicalParam_01^.lrL2			:= 225;(*LREAL*)
		i_pstStMechanicalParam_01^.lrX1			:= 325;(*LREAL*)
		i_pstStMechanicalParam_01^.lrX3			:= 105;(*LREAL*)
		i_pstStMechanicalParam_01^.lrX5			:= 145;(*LREAL*)
		i_pstStMechanicalParam_01^.lrX6			:= 464;(*LREAL*)
		i_pstStMechanicalParam_01^.lrY1			:= 700;(*LREAL*)
		i_pstStMechanicalParam_01^.lrY3			:= 882.5;(*LREAL*)
		i_pstStMechanicalParam_01^.lrY5			:= 1230;(*LREAL*)
		i_pstStMechanicalParam_01^.lrY6			:= 1075;(*LREAL*)
	END_IF
	IF i_pstStMechanicalParam_02<>0 THEN
		i_pstStMechanicalParam_02^.lrD1			:= 100;(**)
		i_pstStMechanicalParam_02^.lrD3			:= 100;(**)
		i_pstStMechanicalParam_02^.lrDR			:= 135;(**)
		i_pstStMechanicalParam_02^.lrX1			:= 325;(**)
		i_pstStMechanicalParam_02^.lrX5			:= 145;(**)
		i_pstStMechanicalParam_02^.lrX6			:= 464;(**)
		i_pstStMechanicalParam_02^.lrY1			:= 700;(**)
		i_pstStMechanicalParam_02^.lrY5			:= 1230;(**)
		i_pstStMechanicalParam_02^.lrY6			:= 1075;(**)
	END_IF
	IF i_pstStMechanicalParam_03<>0 THEN
		i_pstStMechanicalParam_03^.lrD2			:= 100;(**)
		i_pstStMechanicalParam_03^.lrD3			:= 100;(**)
		i_pstStMechanicalParam_03^.lrD4			:= 135;(**)
		i_pstStMechanicalParam_03^.lrD5			:= 100;(**)
		i_pstStMechanicalParam_03^.lrD6			:= 80;(**)
		i_pstStMechanicalParam_03^.lrH12		:= 70;(**)
		i_pstStMechanicalParam_03^.lrM			:= 100;(**)
		i_pstStMechanicalParam_03^.lrN			:= 100;(**)
		i_pstStMechanicalParam_03^.lrX1			:= 325;(**)
		i_pstStMechanicalParam_03^.lrX2			:= 0;(**)
		i_pstStMechanicalParam_03^.lrX3			:= 105;(**)
		i_pstStMechanicalParam_03^.lrX4			:= 640;(**)
		i_pstStMechanicalParam_03^.lrX5			:= 145;(**)
		i_pstStMechanicalParam_03^.lrX6			:= 464;(**)
		i_pstStMechanicalParam_03^.lrY1			:= 700;(**)
		i_pstStMechanicalParam_03^.lrY2			:= 0;(**)
		i_pstStMechanicalParam_03^.lrY3			:= 882.5;(**)
		i_pstStMechanicalParam_03^.lrY4			:= 0;(**)
		i_pstStMechanicalParam_03^.lrY5			:= 1230;(**)
		i_pstStMechanicalParam_03^.lrY6			:= 1075;(**)
	END_IF
	IF i_pstStMechanicalParam_05<>0 THEN
		(*2026.08.27.095847 默认值暂未处理*)
		i_pstStMechanicalParam_05^.rX1:= 167;
		i_pstStMechanicalParam_05^.rX2:= 135;
		i_pstStMechanicalParam_05^.rX3:= 300;
		i_pstStMechanicalParam_05^.rX4:= 454;

		i_pstStMechanicalParam_05^.rY0:= 700;
		i_pstStMechanicalParam_05^.rY1:= 1255;
		i_pstStMechanicalParam_05^.rY4:= 1075;

		i_pstStMechanicalParam_05^.rD1:= 100;
		i_pstStMechanicalParam_05^.rD2:= 100;
		i_pstStMechanicalParam_05^.rD3:= 135;
		i_pstStMechanicalParam_05^.rD4:= 100;

		i_pstStMechanicalParam_05^.rY2:= 1109;(*[AI修改20260829]rL2_3改rY2|辊2安装高度,机台图纸值*)
	END_IF

	iResult:=1;
ELSE
	iResult:=-1;
END_IF

(* ---- KS_RstSysParam_UnSave.st ---- *)
(*@CES
Name=KS_RstSysParam_UnSave
Type=FunctionBlock
TypeGuid=6f9dac99-8de1-4efc-8465-68ac443b7d08
Guid=a7b887dc-87a6-43de-9951-73882ec7d195
HasDeclaration=True
HasImplementation=True
*)
{DECLARATION}
FUNCTION KS_RstSysParam_UnSave : INT
VAR_INPUT
	i_pstStSysParam_UnSave: POINTER TO StSysParam_UnSave;
	i_pstStSysParam_UnSave_RSV: POINTER TO StRSV_SysParam_UnSave;
END_VAR
VAR
	iResult: INT;
END_VAR

{IMPLEMENTATION}
iResult:=0;

IF i_pstStSysParam_UnSave<>0 AND i_pstStSysParam_UnSave_RSV<>0 THEN
	SysMemSet(ADR(i_pstStSysParam_UnSave_RSV^.abyRSV_SysParam_UnSave),
				0,
				SIZEOF(i_pstStSysParam_UnSave_RSV^.abyRSV_SysParam_UnSave));
	i_pstStSysParam_UnSave^.byCurrUsrLevel					:= 0;
	i_pstStSysParam_UnSave^.diEncPos_Virtual                := 65536;
	i_pstStSysParam_UnSave^.xCommEn_Tcp                     := FALSE;
	i_pstStSysParam_UnSave^.xOpenSocketing                  := FALSE;
	i_pstStSysParam_UnSave^.xOpenSocketDne                  := FALSE;
	i_pstStSysParam_UnSave^.xOpenSocketFailed               := FALSE;
	i_pstStSysParam_UnSave^.xConnectOk_Tcp                  := FALSE;
	i_pstStSysParam_UnSave^.byConnectSts_Tcp                := 0;
	SysMemSet(ADR(i_pstStSysParam_UnSave^.abyReserved_Tcp),
				0,
				SIZEOF(i_pstStSysParam_UnSave^.abyReserved_Tcp));

	i_pstStSysParam_UnSave^.xCommEn_WatchDevice_Tcp         := FALSE;
	i_pstStSysParam_UnSave^.xOpenSocketing_WatchDevice      := FALSE;
	i_pstStSysParam_UnSave^.xOpenSocketDne_WatchDevice      := FALSE;
	i_pstStSysParam_UnSave^.xOpenSocketFailed_WatchDevice   := FALSE;
	i_pstStSysParam_UnSave^.xConnectOk_WatchDevice_Tcp      := FALSE;
	i_pstStSysParam_UnSave^.byConnectSts_WatchDevice_Tcp    := 0;
	SysMemSet(ADR(i_pstStSysParam_UnSave^.abyReserved1_Tcp),
				0,
				SIZEOF(i_pstStSysParam_UnSave^.abyReserved1_Tcp));

	i_pstStSysParam_UnSave^.xCommEn_485                     := FALSE;
	i_pstStSysParam_UnSave^.xOpenPortDne                    := FALSE;
	i_pstStSysParam_UnSave^.xOpenPortFailed                 := FALSE;
	i_pstStSysParam_UnSave^.xCommEn_WatchDevice_485         := FALSE;
	i_pstStSysParam_UnSave^.byConnectSts_485                := 0;
	SysMemSet(ADR(i_pstStSysParam_UnSave^.abyReserved_485),
				0,
				SIZEOF(i_pstStSysParam_UnSave^.abyReserved_485));

	i_pstStSysParam_UnSave^.rAO0_WaterValue_Start           := 50;
	i_pstStSysParam_UnSave^.rAO0_WaterValue_Start2          := 80;
(*	i_pstStSysParam_UnSave^.stStSysCfgStruct                := 0;(*系统配置初始化怎么处理*)
	*)
	i_pstStSysParam_UnSave^.byTaperUnitType:= 0;
	i_pstStSysParam_UnSave^.byArcDeCoupleStepTest			:= 0;
	i_pstStSysParam_UnSave^.xSaveFineSampleData_ToArc		:= FALSE;
	i_pstStSysParam_UnSave^.byCurGrpId_HMI					:= 1;
	iResult:=1;
ELSE
	iResult:=-1;
END_IF

(* ---- KS_RstUnitParam_Save.st ---- *)
(*@CES
Name=KS_RstUnitParam_Save
Type=FunctionBlock
TypeGuid=6f9dac99-8de1-4efc-8465-68ac443b7d08
Guid=7648ef96-3be4-4568-b3eb-0b6ef16921e6
HasDeclaration=True
HasImplementation=True
*)
{DECLARATION}
FUNCTION KS_RstUnitParam_Save : INT
VAR_INPUT
	i_pstStSysParam: POINTER TO StSysParam;
	i_pastStUnitParam_Save: POINTER TO ARRAY [1..MAX_UNIT_NUM] OF StUnitParam_Save;
	i_pastStUnitParam_Save_RSV: POINTER TO ARRAY [1..MAX_UNIT_NUM] OF StRSV_UnitParam_Save;
END_VAR
VAR
	iUnit: INT;
	iResult: INT;
END_VAR

{IMPLEMENTATION}
iResult:=0;

IF i_pastStUnitParam_Save<>0 AND i_pastStUnitParam_Save_RSV<>0 THEN
	FOR iUnit:=1 TO MAX_UNIT_NUM BY 1 DO
		SysMemSet(ADR(i_pastStUnitParam_Save_RSV^[iUnit].abyRSV_UnitParam_Save),
					0,
					SIZEOF(i_pastStUnitParam_Save_RSV^[iUnit].abyRSV_UnitParam_Save));
		i_pastStUnitParam_Save^[iUnit].byGrpId											:= 1;
		i_pastStUnitParam_Save^[iUnit].rGirth_BottomRoller                              := 1005.2154;
		i_pastStUnitParam_Save^[iUnit].uiNum_BottomRoller                               := 8;
		i_pastStUnitParam_Save^[iUnit].uiDen_BottomRoller                               := 1;
		i_pastStUnitParam_Save^[iUnit].rGirth_PrnRoller                                 := 500;
		i_pastStUnitParam_Save^[iUnit].uiNum_PrnRoller                                  := 1;
		i_pastStUnitParam_Save^[iUnit].uiDen_PrnRoller                                  := 1;
		i_pastStUnitParam_Save^[iUnit].rGirth_NetRoller                                 := 502.6548;
		i_pastStUnitParam_Save^[iUnit].uiNum_NetRoller                                  := 1;
		i_pastStUnitParam_Save^[iUnit].uiDen_NetRoller                                  := 1;
		i_pastStUnitParam_Save^[iUnit].rLength_Band                                     := 1000;
		i_pastStUnitParam_Save^[iUnit].rErrLength_Band                                  := 0;
		i_pastStUnitParam_Save^[iUnit].rGirth_StrRoller                                 := 500;
		i_pastStUnitParam_Save^[iUnit].uiNum_StrRoller                                  := 1;
		i_pastStUnitParam_Save^[iUnit].uiDen_StrRoller                                  := 1;
		i_pastStUnitParam_Save^[iUnit].rScrewPitch_Horz                                 := 5;
		i_pastStUnitParam_Save^[iUnit].uiNum_Horz                                       := 1;
		i_pastStUnitParam_Save^[iUnit].uiDen_Horz                                       := 1;
		i_pastStUnitParam_Save^[iUnit].lrLimit_Operate_Horz                             := 0;
		i_pastStUnitParam_Save^[iUnit].lrLimit_Driver_Horz                              := 0;
		i_pastStUnitParam_Save^[iUnit].wCtlmod_PrnRoller_Pressure                       := 1;
		i_pastStUnitParam_Save^[iUnit].rScrewPitch_PrnRoller_Pressure                   := 4;
		i_pastStUnitParam_Save^[iUnit].uiNum_PrnRoller_Pressure                         := 40;
		i_pastStUnitParam_Save^[iUnit].uiDen_PrnRoller_Pressure                         := 1;
		i_pastStUnitParam_Save^[iUnit].rScrewPitch_NetRoller_Pressure                   := 2;
		i_pastStUnitParam_Save^[iUnit].uiNum_NetRoller_Pressure                         := 3;
		i_pastStUnitParam_Save^[iUnit].uiDen_NetRoller_Pressure                         := 1;
		i_pastStUnitParam_Save^[iUnit].rScrewPitch_StrRoller_Pressure                   := 2;
		i_pastStUnitParam_Save^[iUnit].uiNum_StrRoller_Pressure                         := 3;
		i_pastStUnitParam_Save^[iUnit].uiDen_StrRoller_Pressure                         := 1;
		i_pastStUnitParam_Save^[iUnit].rMovementHiSpd_PrnRoller_Pressure                := 10;
		i_pastStUnitParam_Save^[iUnit].rMovementHiSpd_NetRoller_Pressure                := 10;
		i_pastStUnitParam_Save^[iUnit].rMovementLoSpd_PrnRoller_Pressure                := 5;
		i_pastStUnitParam_Save^[iUnit].rMovementLoSpd_NetRoller_Pressure                := 5;
		i_pastStUnitParam_Save^[iUnit].rPos_press_dn_PrnRoller_Pressure_M               := 0;
		i_pastStUnitParam_Save^[iUnit].rPos_press_dn_PrnRoller_Pressure_G               := 0;
		i_pastStUnitParam_Save^[iUnit].rPos_press_up_PrnRoller_Pressure_M               := 0;
		i_pastStUnitParam_Save^[iUnit].rPos_press_up_PrnRoller_Pressure_G               := 0;
		i_pastStUnitParam_Save^[iUnit].rPos_load_unload_PrnRoller_Pressure_M            := 0;
		i_pastStUnitParam_Save^[iUnit].rPos_load_unload_PrnRoller_Pressure_G            := 0;
		i_pastStUnitParam_Save^[iUnit].rPos_press_dn_NetRoller_Pressure_M               := 0;
		i_pastStUnitParam_Save^[iUnit].rPos_press_dn_NetRoller_Pressure_G               := 0;
		i_pastStUnitParam_Save^[iUnit].rPos_press_up_NetRoller_Pressure_M               := 0;
		i_pastStUnitParam_Save^[iUnit].rPos_press_up_NetRoller_Pressure_G               := 0;
		i_pastStUnitParam_Save^[iUnit].rPos_load_unload_NetRoller_Pressure_M            := 0;
		i_pastStUnitParam_Save^[iUnit].rPos_load_unload_NetRoller_Pressure_G            := 0;
		i_pastStUnitParam_Save^[iUnit].rPos_press_dn_StrRoller_Pressure_M               := 0;
		i_pastStUnitParam_Save^[iUnit].rPos_press_dn_StrRoller_Pressure_G               := 0;
		i_pastStUnitParam_Save^[iUnit].rPos_press_up_StrRoller_Pressure_M               := 0;
		i_pastStUnitParam_Save^[iUnit].rPos_press_up_StrRoller_Pressure_G               := 0;
		i_pastStUnitParam_Save^[iUnit].rPos_load_unload_StrRoller_Pressure_M            := 0;
		i_pastStUnitParam_Save^[iUnit].rPos_load_unload_StrRoller_Pressure_G            := 0;
		i_pastStUnitParam_Save^[iUnit].rGirth_Confirmed_press_dn_PrnRoller              := 520;
		i_pastStUnitParam_Save^[iUnit].rGirth_Confirmed_press_dn_NetRoller              := 508.94;
		i_pastStUnitParam_Save^[iUnit].rGirth_Confirmed_press_dn_StrRoller              := 500;
//		i_pastStUnitParam_Save^[iUnit].bySts_PrfPosAndEncPosDir                         := 0;
//		i_pastStUnitParam_Save^[iUnit].bySts_PrfPosAndActEncPosDirDir                   := 0;
		i_pastStUnitParam_Save^[iUnit].wFlag_PressFun                                   := 0;
		i_pastStUnitParam_Save^[iUnit].lrAbsEncZeroPos_PrnRoller_Pressure_M             := 0;
		i_pastStUnitParam_Save^[iUnit].lrAbsEncZeroPos_PrnRoller_Pressure_G             := 0;
		i_pastStUnitParam_Save^[iUnit].lrAbsEncZeroPos_NetRoller_Pressure_M             := 0;
		i_pastStUnitParam_Save^[iUnit].lrAbsEncZeroPos_NetRoller_Pressure_G             := 0;
		i_pastStUnitParam_Save^[iUnit].lrAbsEncLimMin_PrnRoller_Pressure_M              := 0;
		i_pastStUnitParam_Save^[iUnit].lrAbsEncLimMax_PrnRoller_Pressure_G              := 0;
		i_pastStUnitParam_Save^[iUnit].lrAbsEncLimMin_NetRoller_Pressure_M              := 0;
		i_pastStUnitParam_Save^[iUnit].lrAbsEncLimMax_NetRoller_Pressure_G              := 0;
		i_pastStUnitParam_Save^[iUnit].xConfirmAbsEncZeroPosDne_PrnRoller_Pressure_M    := FALSE;
		i_pastStUnitParam_Save^[iUnit].xConfirmAbsEncZeroPosDne_PrnRoller_Pressure_G    := FALSE;
		i_pastStUnitParam_Save^[iUnit].xConfirmAbsEncZeroPosDne_NetRoller_Pressure_M    := FALSE;
		i_pastStUnitParam_Save^[iUnit].xConfirmAbsEncZeroPosDne_NetRoller_Pressure_G    := FALSE;
		i_pastStUnitParam_Save^[iUnit].xConfirmload_unloadPosDne_PrnRoller_Pressure_M   := FALSE;
		i_pastStUnitParam_Save^[iUnit].xConfirmload_unloadPosDne_PrnRoller_Pressure_G   := FALSE;
		i_pastStUnitParam_Save^[iUnit].xConfirmload_unloadPosDne_NetRoller_Pressure_M   := FALSE;
		i_pastStUnitParam_Save^[iUnit].xConfirmload_unloadPosDne_NetRoller_Pressure_G   := FALSE;
		i_pastStUnitParam_Save^[iUnit].xConfirmDnPosDne_PrnRoller_Pressure_M            := FALSE;
		i_pastStUnitParam_Save^[iUnit].xConfirmDnPosDne_PrnRoller_Pressure_G            := FALSE;
		i_pastStUnitParam_Save^[iUnit].xConfirmDnPosDne_NetRoller_Pressure_M            := FALSE;
		i_pastStUnitParam_Save^[iUnit].xConfirmDnPosDne_NetRoller_Pressure_G            := FALSE;
		i_pastStUnitParam_Save^[iUnit].xEnable_arc                                      := TRUE;
		IF i_pastStUnitParam_Save^[iUnit].byGrpId<>1 AND i_pastStUnitParam_Save^[iUnit].byGrpId<>2 THEN
			i_pastStUnitParam_Save^[iUnit].byGrpId:= 1;
		END_IF

		i_pastStUnitParam_Save^[iUnit].iMarkTypeId                                      :=
				i_pstStSysParam^.astStGrpParam_Save[i_pastStUnitParam_Save^[iUnit].byGrpId].iMarkTypeId;
		i_pastStUnitParam_Save^[iUnit].iMarkArrangeMode                                 :=
				i_pstStSysParam^.astStGrpParam_Save[i_pastStUnitParam_Save^[iUnit].byGrpId].iMarkArrangeMode;
		i_pastStUnitParam_Save^[iUnit].iGateWidthPhy                                    := 20;
		i_pastStUnitParam_Save^[iUnit].iGateWidthRoundPoints                            := 160;
		i_pastStUnitParam_Save^[iUnit].iGateWidthFinePoints                             := 1000;
		i_pastStUnitParam_Save^[iUnit].iGateSa                                          := 0;
		i_pastStUnitParam_Save^[iUnit].iGateSaEx                                        := 0;
		i_pastStUnitParam_Save^[iUnit].rAlr_V                                           := 0.2;
		i_pastStUnitParam_Save^[iUnit].rAdj_V                                           := 0;
		i_pastStUnitParam_Save^[iUnit].byAvg_V                                          := 3;
		i_pastStUnitParam_Save^[iUnit].iKp_V                                            := 2;
		i_pastStUnitParam_Save^[iUnit].iKi_V                                            := 0;
		i_pastStUnitParam_Save^[iUnit].iKd_V                                            := 0;
		i_pastStUnitParam_Save^[iUnit].rDeadzoneMin_V                                   := 0;
		i_pastStUnitParam_Save^[iUnit].rAlr_H                                           := 0.2;
		i_pastStUnitParam_Save^[iUnit].rAdj_H                                           := 0;
		i_pastStUnitParam_Save^[iUnit].byAvg_H                                          := 3;
		i_pastStUnitParam_Save^[iUnit].iKp_H                                            := 3;
		i_pastStUnitParam_Save^[iUnit].iKi_H                                            := 0;
		i_pastStUnitParam_Save^[iUnit].iKd_H                                            := 8;
		i_pastStUnitParam_Save^[iUnit].rDeadzoneMin_H                                   := 0.01;
		i_pastStUnitParam_Save^[iUnit].rDeadzoneMax_H                                   := 5;
		i_pastStUnitParam_Save^[iUnit].lrPreReg_Length_V                                := 0;
		i_pastStUnitParam_Save^[iUnit].lrFilmLengthFromPrevUnit                         := 7500;
		i_pastStUnitParam_Save^[iUnit].lrPreReg_Adjust                                  := 0;
		i_pastStUnitParam_Save^[iUnit].dwFlag_Ctl                                       := 0;
		i_pastStUnitParam_Save^[iUnit].dwFlag_Sts                                       := 0;
		i_pastStUnitParam_Save^[iUnit].diPreReg_AdjustVal_H                             := 0;
		i_pastStUnitParam_Save^[iUnit].lrAI_med_CoatingPrn                              := 0;
		i_pastStUnitParam_Save^[iUnit].xSwitchOn_CoatingPrn                             := FALSE;
		i_pastStUnitParam_Save^[iUnit].xReverseAdj_CoatingPrn                           := FALSE;
		i_pastStUnitParam_Save^[iUnit].byAdjMode_CoatingPrn                             := 0;
		i_pastStUnitParam_Save^[iUnit].iKp_CoatingPrn                                   := 30;
		i_pastStUnitParam_Save^[iUnit].iKi_CoatingPrn                                   := 30;
		i_pastStUnitParam_Save^[iUnit].iKd_CoatingPrn                                   := 60;
		i_pastStUnitParam_Save^[iUnit].bySensorType_CoatingPrn                          := 0;
		i_pastStUnitParam_Save^[iUnit].lrAI_CoatingPrn                                  := 0;
		i_pastStUnitParam_Save^[iUnit].lrGirth_Using_CoatingPrn                         := 500;
		i_pastStUnitParam_Save^[iUnit].bySignalGain                                     := 0;
		i_pastStUnitParam_Save^[iUnit].xLinkage                                         := FALSE;
		i_pastStUnitParam_Save^[iUnit].rInversedPrecision                               := 0.02;
		i_pastStUnitParam_Save^[iUnit].byCouplingMask                                   := 1;
		i_pastStUnitParam_Save^[iUnit].rHigh_Prn_Roller                                 := 50;
		i_pastStUnitParam_Save^[iUnit].rHigh_Net_Roller                                 := 50;
		i_pastStUnitParam_Save^[iUnit].rweigth_Prn_Bottom_Confirm                       := 0;
		i_pastStUnitParam_Save^[iUnit].rweigth_Prn_Net_Confirm                          := 0;
		i_pastStUnitParam_Save^[iUnit].rweigth_Net_Prn_Confirm                          := 0;
		i_pastStUnitParam_Save^[iUnit].rweigth_Net_Load_Confirm                         := 0;
		i_pastStUnitParam_Save^[iUnit].dwColor_Print                                    := 0;
		i_pastStUnitParam_Save^[iUnit].wLines_Net_Roller                                := 500;
		i_pastStUnitParam_Save^[iUnit].rStep_Pressure_Prn_Net                           := 0;
		i_pastStUnitParam_Save^[iUnit].xConfirmDnPosDne_StrRoller_Pressure_M            := FALSE;
		i_pastStUnitParam_Save^[iUnit].xConfirmDnPosDne_StrRoller_Pressure_G            := FALSE;
		i_pastStUnitParam_Save^[iUnit].lrEncPosPrintDn_Prn_M                            := 0;
		i_pastStUnitParam_Save^[iUnit].lrEncPosPrintDn_Prn_G                            := 0;
		i_pastStUnitParam_Save^[iUnit].lrEncPosPrintDn_Net_M                            := 0;
		i_pastStUnitParam_Save^[iUnit].lrEncPosPrintDn_Net_G                            := 0;
		i_pastStUnitParam_Save^[iUnit].lrEncPosPrintDn_Str_M                            := 0;
		i_pastStUnitParam_Save^[iUnit].lrEncPosPrintDn_Str_G                            := 0;
		i_pastStUnitParam_Save^[iUnit].lrEncPosParallel_Prn_M                           := 0;
		i_pastStUnitParam_Save^[iUnit].lrEncPosParallel_Prn_G                           := 0;
		i_pastStUnitParam_Save^[iUnit].lrEncPosParallel_Net_M                           := 0;
		i_pastStUnitParam_Save^[iUnit].lrEncPosParallel_Net_G                           := 0;
		i_pastStUnitParam_Save^[iUnit].lrEncPosParallel_Str_M                           := 0;
		i_pastStUnitParam_Save^[iUnit].lrEncPosParallel_Str_G                           := 0;
		i_pastStUnitParam_Save^[iUnit].lrPrintPosOffsetDn_Prn_M                         := 0;
		i_pastStUnitParam_Save^[iUnit].lrPrintPosOffsetDn_Prn_G                         := 0;
		i_pastStUnitParam_Save^[iUnit].lrPrintPosOffsetDn_Net_M                         := 0;
		i_pastStUnitParam_Save^[iUnit].lrPrintPosOffsetDn_Net_G                         := 0;
		i_pastStUnitParam_Save^[iUnit].lrPrintPosOffsetDn_Str_M                         := 0;
		i_pastStUnitParam_Save^[iUnit].lrPrintPosOffsetDn_Str_G                         := 0;
//		i_pastStUnitParam_Save^[iUnit].adiEncPos_Start_Virtual_0                        := 0;
		i_pastStUnitParam_Save^[iUnit].diEncPos_Start_Virtual_0                         := 0;
		i_pastStUnitParam_Save^[iUnit].diSampleNum                                      := 1;
		i_pastStUnitParam_Save^[iUnit].diSampleDen                                      := 1;
		i_pastStUnitParam_Save^[iUnit].liABSPos_Prn_M                                   := 0;
		i_pastStUnitParam_Save^[iUnit].liABSPos_Prn_G                                   := 0;
		i_pastStUnitParam_Save^[iUnit].liABSPos_Net_M                                   := 0;
		i_pastStUnitParam_Save^[iUnit].liABSPos_Net_G                                   := 0;
		i_pastStUnitParam_Save^[iUnit].liABSPos_Str_M                                   := 0;
		i_pastStUnitParam_Save^[iUnit].liABSPos_Str_G                                   := 0;
		i_pastStUnitParam_Save^[iUnit].axPressLimit_Min[1]                                 := FALSE;
		i_pastStUnitParam_Save^[iUnit].axPressLimit_Min[2]                                 := FALSE;
		i_pastStUnitParam_Save^[iUnit].axPressLimit_Min[3]                                 := FALSE;
		i_pastStUnitParam_Save^[iUnit].axPressLimit_Max[1]                                 := FALSE;
		i_pastStUnitParam_Save^[iUnit].axPressLimit_Max[2]                                 := FALSE;
		i_pastStUnitParam_Save^[iUnit].axPressLimit_Max[3]                                 := FALSE;
		i_pastStUnitParam_Save^[iUnit].lrEncPosLimit_Prn_M_Max                          := 0;
		i_pastStUnitParam_Save^[iUnit].lrEncPosLimit_Prn_G_Max                          := 0;
		i_pastStUnitParam_Save^[iUnit].lrEncPosLimit_Net_M_Max                          := 0;
		i_pastStUnitParam_Save^[iUnit].lrEncPosLimit_Net_G_Max                          := 0;
		i_pastStUnitParam_Save^[iUnit].lrEncPosLimit_Str_M_Max                          := 0;
		i_pastStUnitParam_Save^[iUnit].lrEncPosLimit_Str_G_Max                          := 0;
		i_pastStUnitParam_Save^[iUnit].rLength_Printing                                 := 1040.68;
		i_pastStUnitParam_Save^[iUnit].iBandLengthFilterCnt                             := 10;
		i_pastStUnitParam_Save^[iUnit].iCoefOfCoupling_V                                := 100;
		i_pastStUnitParam_Save^[iUnit].byFollowColorId                                  := 0;
		i_pastStUnitParam_Save^[iUnit].xWaitFilmLenth_Follow1U                          := FALSE;
		i_pastStUnitParam_Save^[iUnit].wButtonFun_Lamp                                  := 0;
		i_pastStUnitParam_Save^[iUnit].wSwitchFun										:= 0;
//		i_pastStUnitParam_Save^[iUnit].dwSlaveBtn_HMI                                   := 0;
		i_pastStUnitParam_Save^[iUnit].rLong_Step_Roller_Pressure                       := 5;
		i_pastStUnitParam_Save^[iUnit].rShort_Step_Roller_Pressure                      := 0.5;
		i_pastStUnitParam_Save^[iUnit].rSV_UnitTemCtl                                   := 50;
		i_pastStUnitParam_Save^[iUnit].dwCtlBits_UnitBaseCraft                          := 0;
		i_pastStUnitParam_Save^[iUnit].rHz_UnitInkRoller_ManuallySet                    := 20;
		i_pastStUnitParam_Save^[iUnit].rCoeff_UnitInkRoller_Auto                        := 1;

		i_pastStUnitParam_Save^[iUnit].rHz_UnitScraper_ManuallySet                      := 20;
		i_pastStUnitParam_Save^[iUnit].rCoeff_UnitScraper_Auto                          := 1;
		i_pastStUnitParam_Save^[iUnit].rHz_UnitHotWind_ManuallySet                      := 20;
		i_pastStUnitParam_Save^[iUnit].rHz_UnitHotWind_2_ManuallySet                    := 20;
		i_pastStUnitParam_Save^[iUnit].byHotBlower_AO                                   := 20;
		i_pastStUnitParam_Save^[iUnit].wAirReturnWindDoorValue                          := 50;
		i_pastStUnitParam_Save^[iUnit].wAirExhaustWindDoorValue                         := 50;
		i_pastStUnitParam_Save^[iUnit].rHz_UnitExhaust_ManuallySet              		  := 20;

		i_pastStUnitParam_Save^[iUnit].bySignalSelect                                   := 0;
		i_pastStUnitParam_Save^[iUnit].rOffset_T1:=1.73;
		i_pastStUnitParam_Save^[iUnit].rSource_Light_T1:=0.15;
		i_pastStUnitParam_Save^[iUnit].rBias_T1:=2;
		i_pastStUnitParam_Save^[iUnit].rBrightness_Light_T1:=0.15;
		i_pastStUnitParam_Save^[iUnit].rOffset_T2:=1.73;
		i_pastStUnitParam_Save^[iUnit].rSource_Light_T2:=0.15;
		i_pastStUnitParam_Save^[iUnit].rBias_T2:=2;
		i_pastStUnitParam_Save^[iUnit].rBrightness_Light_T2:=0.15;

		i_pastStUnitParam_Save^[iUnit].rK_ArcErr_Lp:= 30;
		i_pastStUnitParam_Save^[iUnit].rFilmLengthFromPrevPressUnit:=8000;(*mm*)

		i_pastStUnitParam_Save^[iUnit].byAve_v_extra:= 3;
		i_pastStUnitParam_Save^[iUnit].xWaitFilmLenth_FollowPreU:= FALSE;
		(*增加参数初始化2025.3.5.161313-套色新算法参数相关*)
		i_pastStUnitParam_Save^[iUnit].stStArc_Mol_Param.xUse_NewArcMol		:= FALSE;
		i_pastStUnitParam_Save^[iUnit].stStArc_Mol_Param.xUsePID_Mol			:= FALSE;
		i_pastStUnitParam_Save^[iUnit].stStArc_Mol_Param.rKadj_PID_Mol		:= 20;
		i_pastStUnitParam_Save^[iUnit].stStArc_Mol_Param.rKadj_I_Mol			:= 1.5;
		i_pastStUnitParam_Save^[iUnit].stStArc_Mol_Param.byKadj_SetType		:= 0;
		i_pastStUnitParam_Save^[iUnit].stStArc_Mol_Param.rKadj_PID_Mol_SteadySts:= 20;
		i_pastStUnitParam_Save^[iUnit].stStArc_Mol_Param.rKadj_I_Mol_SteadySts:= 1;
		i_pastStUnitParam_Save^[iUnit].stStArc_Mol_Param.rMargin_Mag_Arc		:= 20;
		i_pastStUnitParam_Save^[iUnit].stStArc_Mol_Param.rMargin_Phi_Arc		:= 50;

		i_pastStUnitParam_Save^[iUnit].stStArc_Mol_Param.xUseAntiNotch_Arc	:= FALSE;
		i_pastStUnitParam_Save^[iUnit].stStArc_Mol_Param.rWn_Arc				:= 0.08;
		i_pastStUnitParam_Save^[iUnit].stStArc_Mol_Param.rBw_Arc				:= 0.08;
		i_pastStUnitParam_Save^[iUnit].stStArc_Mol_Param.rDp_Arc				:= 10;
		i_pastStUnitParam_Save^[iUnit].stStArc_Mol_Param.xUsePeriodic		:= FALSE;
		i_pastStUnitParam_Save^[iUnit].stStArc_Mol_Param.rG_Periodic			:= 0.5;
		i_pastStUnitParam_Save^[iUnit].stStArc_Mol_Param.rW_Periodic			:= 2;
		i_pastStUnitParam_Save^[iUnit].stStArc_Mol_Param.stStArcSpeedUpParam.rK:= 1;
		i_pastStUnitParam_Save^[iUnit].stStArc_Mol_Param.stStArcSpeedUpParam.rA2:= 40;
		i_pastStUnitParam_Save^[iUnit].stStArc_Mol_Param.stStArcSpeedUpParam.rA1:= 6;
		i_pastStUnitParam_Save^[iUnit].stStArc_Mol_Param.stStArcSpeedUpParam.rA0:= 0.01;
		i_pastStUnitParam_Save^[iUnit].stStArc_Mol_Param.stStArcSpeedUpFeedforward.rK:= 2000;
		i_pastStUnitParam_Save^[iUnit].stStArc_Mol_Param.stStArcSpeedUpFeedforward.rK_2:= 2000;

		i_pastStUnitParam_Save^[iUnit].stStArc_Mol_Param.rKp_GC:= 16;
		i_pastStUnitParam_Save^[iUnit].stStArc_Mol_Param.rKi_GC:= 15;
		i_pastStUnitParam_Save^[iUnit].stStArc_Mol_Param.rKd_GC:=0;
		i_pastStUnitParam_Save^[iUnit].stStArc_Mol_Param.rN_GC:= 0;
		i_pastStUnitParam_Save^[iUnit].stStArc_Mol_Param.xCompensateEn_H:=FALSE;
		i_pastStUnitParam_Save^[iUnit].stStArc_Mol_Param.byCompensateValue_Hor:=50;(*丝*)
		i_pastStUnitParam_Save^[iUnit].stStArc_Mol_Param.byMaxAddValue_Total_Hor:=5;(*mm*)

			(*新增变量|wang.nt|2025.08.07.204018*)
		i_pastStUnitParam_Save^[iUnit].rStep_OfChangeGirth 					:= 0.01;  (*涂布版轴修改步幅*)
		i_pastStUnitParam_Save^[iUnit].uiTimeMs_RollerPressUpKeep 			:= 0;      (*压辊双气缸-离压保持时间*)
		//9905界面内容
		i_pastStUnitParam_Save^[iUnit].rAxisVelPrf_Coeff1 					:= -200	;
		i_pastStUnitParam_Save^[iUnit].rAxisVelPrf_Coeff2 					:= 0.03	;
		i_pastStUnitParam_Save^[iUnit].rAxisVelPrf_Coeff3 					:= 1	;
		i_pastStUnitParam_Save^[iUnit].rMargin_Mag_Arc 						:= 20	;
		i_pastStUnitParam_Save^[iUnit].rMargin_Phi_Arc 						:= 50	;
		i_pastStUnitParam_Save^[iUnit].rKp_MolCal 							:= 16	;
		i_pastStUnitParam_Save^[iUnit].rKi_MolCal 							:= 8	;
		i_pastStUnitParam_Save^[iUnit].rFilmLengthFromPrevPressUnit 		:= 8000	;
		i_pastStUnitParam_Save^[iUnit].byCompensateValue_Hor 				:= 50	;
		i_pastStUnitParam_Save^[iUnit].byMaxAddValue_Total_Hor 				:= 5	;
		i_pastStUnitParam_Save^[iUnit].rWn_Arc 								:= 0.08	;
		i_pastStUnitParam_Save^[iUnit].rBw_Arc 								:= 0.08	;
		i_pastStUnitParam_Save^[iUnit].rDp_Arc 								:= 10	;
		i_pastStUnitParam_Save^[iUnit].rK 									:= 1	;
		i_pastStUnitParam_Save^[iUnit].rA2 									:= 40	;
		i_pastStUnitParam_Save^[iUnit].rA1 									:= 6	;
		i_pastStUnitParam_Save^[iUnit].rA0 									:= 0.01	;
		i_pastStUnitParam_Save^[iUnit].rG_Periodic 							:= 0.5 	;
		i_pastStUnitParam_Save^[iUnit].rW_Periodic 							:= 2	;
		(*2025.8.13.144044增加*)
		i_pastStUnitParam_Save^[iUnit].xFlag_InkRollerRisen:= FALSE;(*2018.7.28.101609\递墨辊升起标志|*)
		i_pastStUnitParam_Save^[iUnit].lrPreReg_ConstVal                          := 6000;
		(*2026.02.28.134214 超旭照明默认开 Hou.N*)
		i_pastStUnitParam_Save^[iUnit].wButtonAndSwitch_ChaoXu.4                          := TRUE;
	END_FOR
	iResult:=1;
ELSE
	iResult:=-1;
END_IF
